// TIA Portal V21 export
FUNCTION_BLOCK "GraphQualification"   // FB, GRAPH
// stored: AutoNumber true
   VAR_INPUT
      ACK_EF : Bool;
      StartCommand : Bool;
      ResetCommand : Bool;
      GuardClosed : Bool;
      SupervisionTrip : Bool;
   END_VAR
   VAR_OUTPUT
      MotorA : Bool;
      MotorB : Bool;
   END_VAR
BEGIN
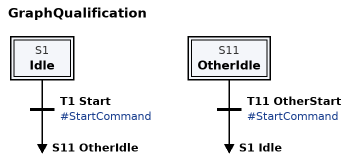
   // sequencer 1: Parallel cycle / Paralleler Ablauf
   INITIAL_STEP Idle:   // S1
      interlock C := #GuardClosed;
      supervision V := #SupervisionTrip;
   END_STEP
   TRANSITION Start FROM Idle TO OtherIdle   // T1, jump
      := #StartCommand;
   END_TRANSITION

   // sequencer 2: Parallel cycle / Paralleler Ablauf
   INITIAL_STEP OtherIdle:   // S11
      interlock C := #GuardClosed;
      supervision V := #SupervisionTrip;
   END_STEP
   TRANSITION OtherStart FROM OtherIdle TO Idle   // T11, jump
      := #StartCommand;
   END_TRANSITION
END_FUNCTION_BLOCK
